INTERFACE I_LimitRule EXTENDS I_Module

PROPERTY Basis : E_LimitBasis
GET
END_GET
END_PROPERTY

METHOD M_Evaluate : ST_LimitOut
VAR_INPUT
	i_stView	: ST_GroupView;
END_VAR
END_METHOD

END_INTERFACE

(* stored: Version 1.1.0.1, ProductVersion 3.1.4024.15
   Itf I_LimitRule: Id {d84dd1d2-3765-40db-b311-784681c8bb38}
   Property Basis: Id {7e2e51b1-be04-4b42-8fc9-efb5dd7a9906}
   Get Get: Id {f2074f08-94cc-4dfa-a33f-1fe1209e96a3}
   Method M_Evaluate: Id {52682d66-04cd-4425-827f-c4a657b815a7} *)
